TYPE ST_EL3351CoeReadData :
STRUCT
	wIdx: WORD;
	bySubIdx: BYTE;
	bReadOK: BOOL;
	nData: UDINT;
	nSize: UDINT;
END_STRUCT
END_TYPE

(* stored: Version 1.1.0.1, ProductVersion 3.1.4024.15
   DUT ST_EL3351CoeReadData: Id {d569db15-bcfd-4082-83e2-69943affb570} *)
